// TIA Portal V15.1 export
// export: Created 2026-11-01T20:56:24.8924892Z, ExportSetting WithDefaults, DisplayName Totally Integrated Automation Portal, DisplayVersion V15.1, DisplayName TIA Portal Openness, DisplayVersion V15.1, DisplayName STEP 7 Professional, DisplayVersion V15.1, DisplayName WinCC Professional, DisplayVersion V15.1
Screen "Screen_1"  480x272, Number=1
  ScreenLayer 
    IOField "I/O field_1" at 16,17 size 96x32  DataFormat=Decimal, FormatPattern=s99999, Mode=InOutput
      ProcessValue := Par_SP
